// TIA Portal V19 export
TYPE "ST_ROBOT"
   STRUCT
      SEND : Struct   // PLC -> ROBOT
         USER_BITS : "ST_USER_BITS_SEND";
         EXTERNALSTART : Bool;
         EXTERNALHOLD : Bool;
         CALLMASTERJOB : Bool;
         ALARMRESET : Bool;
         EXTERNALSERVOON : Bool;
         REDUCESPEED : Bool;
         EDITLOCK : Bool;
         LOWAIRPRESSURE : Bool;
         BUZZER : Bool;
         WATCHDOG : Bool;
         MACHINELOCK : Bool;
         "NOT-USED" : Bool;
         CMD : Int;   // I10
         CMD_ID : Int;   // I11
         X : Int;   // I12 (X, mm)
         Y : Int;   // I13 (Y, mm)
         Z : Int;   // I14 (Z, mm)
         Rx : Int;
         Ry : Int;
         Rz : Int;
         PARAM_1 : Int;
         PARAM_2 : Int;
         PARAM_3 : Int;
         PARAM_4 : Int;
         PARAM_5 : Int;
         PARAM_6 : Int;
         PARAM_7 : Int;
         PARAM_8 : Int;
         PARAM_9 : Int;
         FUNCTION_ID : Int;   // Debug only, not send to the robot Additional system signals from the supplied mapping.
         INVALIDCOLLISIONDETECT : Bool;   // SEND byte 1, bit 3
         CONTINUOUSCYCLESELECT : Bool;   // SEND byte 1, bit 4
         ONECYCLESELECT : Bool;   // SEND byte 1, bit 5
         AUTOBACKUP : Bool;   // SEND byte 1, bit 7
         WORKPROHIBIT_R1 : Bool;   // SEND byte 2, bit 0
         WORKPROHIBIT_R2 : Bool;   // SEND byte 2, bit 1
         WORKPROHIBIT_R3 : Bool;   // SEND byte 2, bit 2
         WORKPROHIBIT_R4 : Bool;   // SEND byte 2, bit 3
         WORKPROHIBIT_R5 : Bool;   // SEND byte 2, bit 4
         WORKPROHIBIT_R6 : Bool;   // SEND byte 2, bit 5
         WORKPROHIBIT_R7 : Bool;   // SEND byte 2, bit 6
         WORKPROHIBIT_R8 : Bool;   // SEND byte 2, bit 7
         SEQUENCEWAIT_R1 : Bool;   // SEND byte 3, bit 0
         SEQUENCEWAIT_R2 : Bool;   // SEND byte 3, bit 1
         SEQUENCEWAIT_R3 : Bool;   // SEND byte 3, bit 2
         SEQUENCEWAIT_R4 : Bool;   // SEND byte 3, bit 3
         SEQUENCEWAIT_R5 : Bool;   // SEND byte 3, bit 4
         SEQUENCEWAIT_R6 : Bool;   // SEND byte 3, bit 5
         SEQUENCEWAIT_R7 : Bool;   // SEND byte 3, bit 6
         SEQUENCEWAIT_R8 : Bool;   // SEND byte 3, bit 7
         SEQUENCEWAIT_S1 : Bool;   // SEND byte 4, bit 0
         SEQUENCEWAIT_S2 : Bool;   // SEND byte 4, bit 1
         SEQUENCEWAIT_S3 : Bool;   // SEND byte 4, bit 2
         SEQUENCEWAIT_S4 : Bool;   // SEND byte 4, bit 3
         SEQUENCEWAIT_S5 : Bool;   // SEND byte 4, bit 4
         SEQUENCEWAIT_S6 : Bool;   // SEND byte 4, bit 5
         SEQUENCEWAIT_S7 : Bool;   // SEND byte 4, bit 6
         SEQUENCEWAIT_S8 : Bool;   // SEND byte 4, bit 7
         STEPBACK_R1 : Bool;   // SEND byte 5, bit 0
         STEPBACK_R2 : Bool;   // SEND byte 5, bit 1
         STEPBACK_R3 : Bool;   // SEND byte 5, bit 2
         STEPBACK_R4 : Bool;   // SEND byte 5, bit 3
         STEPBACK_R5 : Bool;   // SEND byte 5, bit 4
         STEPBACK_R6 : Bool;   // SEND byte 5, bit 5
         STEPBACK_R7 : Bool;   // SEND byte 5, bit 6
         STEPBACK_R8 : Bool;   // SEND byte 5, bit 7
         PARAM_10 : Int;
         PARAM_11 : Int;
         PARAM_12 : Int;
         PARAM_13 : Int;   // Retained for compatibility; not transmitted in this layout.
         PARAM_BYTE_62 : Byte;   // Byte 62 only; one-byte parameter (0..255).
      END_STRUCT;
      RECEIVE : Struct   // ROBOT -> PLC
         USER_BITS : "ST_USER_BITS_RECIEVE";
         RUNNING : Bool;
         SERVOISON : Bool;
         TOPMASTERJOB : Bool;
         ALARM : Bool;
         HOLD : Bool;
         REMOTEMODE : Bool;
         PLAYMODE : Bool;
         TEACHMODE : Bool;
         ROBOTCOLLISION : Bool;
         REDUCEDSPEED : Bool;
         "NOT-USED" : Bool;
         ACT_CMDID : Int;
         ACT_X : Int;   // mm
         ACT_Y : Int;   // mm
         ACT_Z : Int;   // mm
         ACT_Rz : Int;
         PARAM_1 : Int;
         PARAM_2 : Int;
         PARAM_3 : Int;
         PARAM_4 : Int;
         PARAM_5 : Int;
         PARAM_6 : Int;
         PARAM_7 : Int;
         PARAM_8 : Int;
         PARAM_9 : Int;   // Additional system signals from the supplied mapping.
         BATTERYALARM : Bool;   // RECEIVE byte 1, bit 0
         WATCHDOG : Bool;   // RECEIVE byte 1, bit 1
         CONTINUOUSCYCLESELECT : Bool;   // RECEIVE byte 1, bit 4
         ONECYCLESELECT : Bool;   // RECEIVE byte 1, bit 5
         DIALOGDISPLAYATSTART : Bool;   // RECEIVE byte 1, bit 6
         ENERGYSAVING : Bool;   // RECEIVE byte 1, bit 7
         MAJORALARM : Bool;   // RECEIVE byte 2, bit 0
         MINORALARM : Bool;   // RECEIVE byte 2, bit 1
         SYSTEMALARM : Bool;   // RECEIVE byte 2, bit 2
         USERALARM : Bool;   // RECEIVE byte 2, bit 3
         SAFETYPLUGINPUT : Bool;   // RECEIVE byte 2, bit 4
         EXTERNALEMERGENCYSTOP : Bool;   // RECEIVE byte 2, bit 5
         TEACHBOXEMERGENCYSTOP : Bool;   // RECEIVE byte 2, bit 6
         EXTERNALHOLD : Bool;   // RECEIVE byte 2, bit 7
         SHOCKDETECTION_R1 : Bool;   // RECEIVE byte 3, bit 0
         SHOCKDETECTION_R2 : Bool;   // RECEIVE byte 3, bit 1
         SHOCKDETECTION_R3 : Bool;   // RECEIVE byte 3, bit 2
         SHOCKDETECTION_R4 : Bool;   // RECEIVE byte 3, bit 3
         SHOCKDETECTION_R5 : Bool;   // RECEIVE byte 3, bit 4
         SHOCKDETECTION_R6 : Bool;   // RECEIVE byte 3, bit 5
         SHOCKDETECTION_R7 : Bool;   // RECEIVE byte 3, bit 6
         SHOCKDETECTION_R8 : Bool;   // RECEIVE byte 3, bit 7
         INCUBE_1 : Bool;   // RECEIVE byte 4, bit 0
         INCUBE_2 : Bool;   // RECEIVE byte 4, bit 1
         INCUBE_3 : Bool;   // RECEIVE byte 4, bit 2
         INCUBE_4 : Bool;   // RECEIVE byte 4, bit 3
         INCUBE_5 : Bool;   // RECEIVE byte 4, bit 4
         INCUBE_6 : Bool;   // RECEIVE byte 4, bit 5
         INCUBE_7 : Bool;   // RECEIVE byte 4, bit 6
         INCUBE_8 : Bool;   // RECEIVE byte 4, bit 7
         INCUBE_9 : Bool;   // RECEIVE byte 5, bit 0
         INCUBE_10 : Bool;   // RECEIVE byte 5, bit 1
         INCUBE_11 : Bool;   // RECEIVE byte 5, bit 2
         INCUBE_12 : Bool;   // RECEIVE byte 5, bit 3
         INCUBE_13 : Bool;   // RECEIVE byte 5, bit 4
         INCUBE_14 : Bool;   // RECEIVE byte 5, bit 5
         INCUBE_15 : Bool;   // RECEIVE byte 5, bit 6
         INCUBE_16 : Bool;   // RECEIVE byte 5, bit 7
         PARAM_10 : Int;
         PARAM_11 : Int;
         PARAM_12 : Int;
         PARAM_13 : Int;
         PARAM_14 : Int;   // Retained for compatibility; not transmitted in this layout.
         PARAM_BYTE_62 : Byte;   // Byte 62 only; one-byte parameter (0..255).
      END_STRUCT;
   END_STRUCT;
END_TYPE
